(* IEC 61131-3 sources: s7-to-codesys/s7conv/tests/snapshots/fixtures/src/POUs/FB_Motor, 2 files *)

(* ---- FB_Motor.decl.st ---- *)
// Назначение: Motor with feedback supervision
//             Пуск по фронту команды, контроль обратной связи через FeedbackTime.
// Автор:      Engineer (исходный блок S7); перевод в ST — s7conv 0.1.0
// Версия:     1.2 (исходный блок S7)
// Документ:   docs/CONVERSION_REPORT.md, docs/MAPPING.md
// Источник:   s7conv/tests/fixtures/motor.scl, строки 14–101, FUNCTION_BLOCK "FB_Motor", FAMILY Drives
// Сгенерировано s7conv: пометки MIGRATION-CHECK и MIGRATION-TODO требуют ручного разбора.
// MIGRATION-CHECK: VAR RETAIN в ФБ: в CODESYS при RETAIN-переменной в retain-памяти хранится весь экземпляр ФБ, в
//                  S7 — только эти переменные (сверить с источником) (стр. 46)
FUNCTION_BLOCK FB_Motor
VAR_INPUT
    cmd : UDT_MotorCmd;
    feedback : BOOL;  // контактор включён
    feedbackTime : TIME := T#3S;
END_VAR
VAR_OUTPUT
    run : BOOL;
    fault : BOOL;
    runTime : TIME;
END_VAR
VAR_IN_OUT
    ack : BOOL;
END_VAR
VAR
    startEdge : R_TRIG;
    fbTimer : TON;
    starts : DINT;
    stat : ST_FB_Motor_stat;
END_VAR
VAR RETAIN
    operatingHours : REAL;
END_VAR
VAR_TEMP
    i : INT;
END_VAR
VAR CONSTANT
    MAX_STARTS : DINT := 1000;
END_VAR

(* ---- FB_Motor.impl.st ---- *)
// REGION Edge detection
startEdge(CLK := cmd.start);
// END_REGION Edge detection

// REGION Mode handling
CASE cmd.mode OF
    0:
        // выведен из работы
        run := FALSE;
    1, 2:
        IF startEdge.Q AND NOT fault THEN
            run := TRUE;
            starts := starts + 1;
        ELSIF cmd.stop THEN
            run := FALSE;
        END_IF
ELSE
    run := FALSE;
END_CASE
// END_REGION Mode handling

// Контроль обратной связи
fbTimer(IN := run AND NOT feedback, PT := feedbackTime, ET => runTime);
IF fbTimer.Q THEN
    fault := TRUE;
    run := FALSE;
END_IF
IF ack THEN
    fault := FALSE;
    ack := FALSE;
END_IF

FOR i := 3 TO 1 BY -1 DO
    stat.history[i] := stat.history[i - 1];
END_FOR
stat.history[0] := run;
stat.lastMode := cmd.mode;
IF starts > MAX_STARTS THEN
    starts := 0;
END_IF
